Staubli VAL3: ifString.pgx

public program ifString(string x_sKey, num x_nIndex, string& x_sMsg)
  local num l_i
  local num l_nSigIndex
  local num l_nSigType
  local num l_nValue
  local bool l_bANDOR1
  local bool l_bANDOR2
  local string l_sMsg1
  local string l_sMsg2
  local string l_sMsg3
  local string l_sANDOR1
  local string l_sANDOR2
begin
  l_sMsg1=""
  l_sMsg2=""
  l_sMsg3=""
  l_nSigType=progTemp:pProgItem[x_sKey].pProgTemplate[x_nIndex].iIfItem.nSigType[0]
  l_nSigIndex=progTemp:pProgItem[x_sKey].pProgTemplate[x_nIndex].iIfItem.nSigIndex[0]
  l_nValue=progTemp:pProgItem[x_sKey].pProgTemplate[x_nIndex].iIfItem.nValue[0]
  if l_nSigType>0 and l_nSigIndex>0
    switch l_nSigType
      case 1
        if l_nValue!=0
          l_sMsg1="DIN"+toString("",l_nSigIndex)+"=true"
        else
          l_sMsg1="DIN"+toString("",l_nSigIndex)+"=false"
        endIf
      break
      case 2
        if l_nValue!=0
          l_sMsg1="DOUT"+toString("",l_nSigIndex)+"=true"
        else
          l_sMsg1="DOUT"+toString("",l_nSigIndex)+"=false"
        endIf
      break
      case 3
        l_sMsg1="AIN"+toString("",l_nSigIndex)+"="+toString("",l_nValue)
      break
      case 4
        l_sMsg1="AOUT"+toString("",l_nSigIndex)+"="+toString("",l_nValue)
      break
    endSwitch
  endIf
  l_bANDOR1=progTemp:pProgItem[x_sKey].pProgTemplate[x_nIndex].iIfItem.bANDOR[0]
  if !l_bANDOR1
    l_sANDOR1=" and "
  else
    l_sANDOR1=" or "
  endIf
  l_bANDOR2=progTemp:pProgItem[x_sKey].pProgTemplate[x_nIndex].iIfItem.bANDOR[1]
  if !l_bANDOR2
    l_sANDOR2=" and "
  else
    l_sANDOR2=" or "
  endIf
  l_nSigType=progTemp:pProgItem[x_sKey].pProgTemplate[x_nIndex].iIfItem.nSigType[1]
  l_nSigIndex=progTemp:pProgItem[x_sKey].pProgTemplate[x_nIndex].iIfItem.nSigIndex[1]
  l_nValue=progTemp:pProgItem[x_sKey].pProgTemplate[x_nIndex].iIfItem.nValue[1]
  if l_nSigType>0 and l_nSigIndex>0

    switch l_nSigType
      case 1
        if l_nValue!=0
          l_sMsg2="DIN"+toString("",l_nSigIndex)+"=true"
        else
          l_sMsg2="DIN"+toString("",l_nSigIndex)+"=false"
        endIf
      break
      case 2
        if l_nValue!=0
          l_sMsg2="DOUT"+toString("",l_nSigIndex)+"=true"
        else
          l_sMsg2="DOUT"+toString("",l_nSigIndex)+"=false"
        endIf
      break
      case 3
        l_sMsg2="AIN"+toString("",l_nSigIndex)+"="+toString("",l_nValue)
      break
      case 4
        l_sMsg2="AOUT"+toString("",l_nSigIndex)+"="+toString("",l_nValue)
      break
    endSwitch
    l_sMsg2=l_sANDOR1+l_sMsg2
  endIf
  l_nSigType=progTemp:pProgItem[x_sKey].pProgTemplate[x_nIndex].iIfItem.nSigType[2]
  l_nSigIndex=progTemp:pProgItem[x_sKey].pProgTemplate[x_nIndex].iIfItem.nSigIndex[2]
  l_nValue=progTemp:pProgItem[x_sKey].pProgTemplate[x_nIndex].iIfItem.nValue[2]
  if l_nSigType>0 and l_nSigIndex>0
    switch l_nSigType
      case 1
        if l_nValue!=0
          l_sMsg3="DIN"+toString("",l_nSigIndex)+"=true"
        else
          l_sMsg3="DIN"+toString("",l_nSigIndex)+"=false"
        endIf
      break
      case 2
        if l_nValue!=0
          l_sMsg3="DOUT"+toString("",l_nSigIndex)+"=true"
        else
          l_sMsg3="DOUT"+toString("",l_nSigIndex)+"=false"
        endIf
      break
      case 3
        l_sMsg3="AIN"+toString("",l_nSigIndex)+"="+toString("",l_nValue)
      break
      case 4
        l_sMsg3="AOUT"+toString("",l_nSigIndex)+"="+toString("",l_nValue)
      break
    endSwitch
    l_sMsg3=l_sANDOR2+l_sMsg3
  endIf

  x_sMsg=l_sMsg1+l_sMsg2+l_sMsg3
end
